(*
SPDX-FileCopyrightText: c 2026 Oleksandr Tiutyk <trofimich@gmail.com>
SPDX-License-Identifier: MIT
License: https://opensource.org/license/mit
*)

(*!
<summary>Checks generic lookup with independent borrowed query values.</summary>
<description>
Owns an inline queue and its copied entry payloads. Run from one task at a stable address.
Teardown clears surviving entries before publication, including after an aborted case.
</description>
*)

{attribute 'no_assign'}
{attribute 'no_explicit_call' := 'do not call this function block directly'}
FUNCTION_BLOCK StaticQueueContainsGenericTest EXTENDS TOF_Testing.SingleCycleTest
VAR_STAT
	{attribute 'hide'}
	_ClassName : STRING := __POUNAME();
END_VAR
VAR
	_Queue : TOF_Collections.Queue<3>(valueValidator := 0);
END_VAR

(*!
<summary>Checks generic lookup with independent borrowed query values.</summary>
*)
METHOD PROTECTED ExecuteTest
VAR
	values : ARRAY [1..4] OF INT := [11, 22, 33, 44];
	query : TOF_Core.GENERIC_VALUE;
END_VAR
_Queue
	.EnqueueCopy(value := values[1])
	.EnqueueCopy(value := values[2])
	.EnqueueCopy(value := values[3]);

query := TOF_Core.GenericValueFactory.FromIntReference(value := values[1]);
Assert.ThatBool(
	actual := _Queue.ContainsGeneric(value := query, releaseValue := FALSE),
	message := "Generic lookup must find the head"
).IsTrue();

query := TOF_Core.GenericValueFactory.FromIntReference(value := values[3]);
Assert.ThatBool(
	actual := _Queue.ContainsGeneric(value := query, releaseValue := FALSE),
	message := "Generic lookup must find the tail"
).IsTrue();

query := TOF_Core.GenericValueFactory.FromIntReference(value := values[4]);
Assert.ThatBool(
	actual := _Queue.ContainsGeneric(value := query, releaseValue := FALSE),
	message := "Generic lookup must report a missing value"
).IsFalse();

Assert.ThatDInt(
	actual := _Queue.Length,
	message := "Generic lookup must preserve queue length"
).ToBe(expected := DINT#3);
END_METHOD

(*!
<summary>Restores the fixture before the runner publishes the result.</summary>
<description>
Also runs after an unexpected exception interrupts the case.
</description>
*)
METHOD PROTECTED AfterTest
_Queue.Clear();
END_METHOD

//! <summary>Borrows the concrete class name. Callers must not modify it.</summary>
{attribute 'monitoring' := 'call'}
PROPERTY ClassName : REFERENCE TO STRING
GET
ClassName REF= _ClassName;
END_GET
END_PROPERTY

//! <summary>Borrows the compiler-initialized namespace name. Callers must not modify it.</summary>
{attribute 'monitoring' := 'call'}
PROPERTY NamespaceName : REFERENCE TO STRING
GET
NamespaceName REF= CurrentNamespace.Name;
END_GET
END_PROPERTY

//! <summary>Reports the concrete instance size in bytes.</summary>
{attribute 'monitoring' := 'call'}
PROPERTY SelfSize : ULINT
GET
SelfSize := XSIZEOF(THIS^);
END_GET
END_PROPERTY

END_FUNCTION_BLOCK

(* stored: Version 1.1.0.1
   POU StaticQueueContainsGenericTest: Id {c9b4bfa2-5d00-407e-baa7-45e6643577cf}, SpecialFunc None
   Method ExecuteTest: Id {0eaf32ad-d092-4556-9b9e-18aa92117da7}
   Method AfterTest: Id {54fdcb61-d812-4364-9601-40d54ab8e99d}
   Property ClassName: Id {a59aa705-657f-48d8-9e2b-01c763657ccc}
   Get Get: Id {1566c06a-5ded-4574-becc-cfe81b0b62f9}
   Property NamespaceName: Id {a142418c-1db4-475f-8064-fdb2631afdee}
   Get Get: Id {ea01f45a-56af-444f-b9eb-cdfb5966cf3b}
   Property SelfSize: Id {c54e5186-b72f-4dac-90f2-14f5cad553a5}
   Get Get: Id {f0562dbd-aa3a-4fd1-a380-bb85332e59ec} *)
